// TIA Portal V20 export
Screen "Pop-up_PN_DEV_DIAG_Counter_Popup"  290x322
  ScreenItem "Background" at 0,0 size 290x322  Type=HmiRectangle
  ScreenItem "Text_ReadedDEVNumbers" at 8,163 size 276x25  Type=HmiTextBox
  ScreenItem "Text_Configured" at 10,37 size 130x25  Type=HmiTextBox
  ScreenItem "Counter_Configured" at 145,38 size 44x23  Type=HmiIOField
  ScreenItem "Text_Faulty" at 10,112 size 130x25  Type=HmiTextBox
  ScreenItem "Counter_Faulty" at 145,113 size 44x23  Type=HmiIOField
  ScreenItem "Text_Deaktivated" at 10,87 size 130x25  Type=HmiTextBox
  ScreenItem "Counter_Deaktivated" at 145,88 size 44x23  Type=HmiIOField
  ScreenItem "Text_Present" at 10,62 size 130x25  Type=HmiTextBox
  ScreenItem "Counter_Present" at 145,63 size 44x23  Type=HmiIOField
  ScreenItem "Text_Problem" at 10,137 size 130x25  Type=HmiTextBox
  ScreenItem "Counter_Problem" at 145,138 size 44x23  Type=HmiIOField
  ScreenItem "Text_MaxDevices" at 10,266 size 130x25  Type=HmiTextBox
  ScreenItem "Text_MaxModules" at 10,291 size 130x25  Type=HmiTextBox
  ScreenItem "Counter_MaxDevices" at 145,267 size 44x23  Type=HmiIOField
  ScreenItem "Counter_Max_Modules" at 145,292 size 44x23  Type=HmiIOField
  ScreenItem "Text_PNDEVCounter" at 1,3 size 288x30  Type=HmiTextBox
  ScreenItem "Text_PLCSettings" at 10,241 size 276x25  Type=HmiTextBox
  ScreenItem "Text_Lowest" at 10,185 size 130x25  Type=HmiTextBox
  ScreenItem "Text_Highest" at 10,210 size 130x25  Type=HmiTextBox
  ScreenItem "Counter_LowDevice" at 145,187 size 44x23  Type=HmiIOField
  ScreenItem "Counter_HighDevice" at 145,212 size 44x23  Type=HmiIOField
  ScreenItem "Cancel Mode_1" at 206,278 size 82x42  Type=HmiButton
  ScreenItem "Background_1" at 8,8 size 290x322  Type=HmiRectangle
  ScreenItem "Text_ReadedDEVNumbers_1" at 16,171 size 276x25  Type=HmiTextBox
  ScreenItem "Text_Configured_1" at 18,45 size 130x25  Type=HmiTextBox
  ScreenItem "Counter_Configured_1" at 153,46 size 44x23  Type=HmiIOField
  ScreenItem "Text_Faulty_1" at 18,120 size 130x25  Type=HmiTextBox
  ScreenItem "Counter_Faulty_1" at 153,121 size 44x23  Type=HmiIOField
  ScreenItem "Text_Deaktivated_1" at 18,95 size 130x25  Type=HmiTextBox
  ScreenItem "Counter_Deaktivated_1" at 153,96 size 44x23  Type=HmiIOField
  ScreenItem "Text_Present_1" at 18,70 size 130x25  Type=HmiTextBox
  ScreenItem "Counter_Present_1" at 153,71 size 44x23  Type=HmiIOField
  ScreenItem "Text_Problem_1" at 18,145 size 130x25  Type=HmiTextBox
  ScreenItem "Counter_Problem_1" at 153,146 size 44x23  Type=HmiIOField
  ScreenItem "Text_MaxDevices_1" at 18,274 size 130x25  Type=HmiTextBox
  ScreenItem "Text_MaxModules_1" at 18,299 size 130x25  Type=HmiTextBox
  ScreenItem "Counter_MaxDevices_1" at 153,275 size 44x23  Type=HmiIOField
  ScreenItem "Counter_Max_Modules_1" at 153,300 size 44x23  Type=HmiIOField
  ScreenItem "Text_PNDEVCounter_1" at 9,11 size 288x30  Type=HmiTextBox
  ScreenItem "Text_PLCSettings_1" at 18,249 size 276x25  Type=HmiTextBox
  ScreenItem "Text_Lowest_1" at 18,193 size 130x25  Type=HmiTextBox
  ScreenItem "Text_Highest_1" at 18,218 size 130x25  Type=HmiTextBox
  ScreenItem "Counter_LowDevice_1" at 153,195 size 44x23  Type=HmiIOField
  ScreenItem "Counter_HighDevice_1" at 153,220 size 44x23  Type=HmiIOField
  ScreenItem "Cancel Mode_2" at 214,286 size 82x42  Type=HmiButton
  ScreenItem "Background_2" at 402,11 size 290x322  Type=HmiRectangle
  ScreenItem "Text_ReadedDEVNumbers_2" at 410,174 size 276x25  Type=HmiTextBox
  ScreenItem "Text_Configured_2" at 412,48 size 130x25  Type=HmiTextBox
  ScreenItem "Counter_Configured_2" at 547,49 size 44x23  Type=HmiIOField
  ScreenItem "Text_Faulty_2" at 412,123 size 130x25  Type=HmiTextBox
  ScreenItem "Counter_Faulty_2" at 547,124 size 44x23  Type=HmiIOField
  ScreenItem "Text_Deaktivated_2" at 412,98 size 130x25  Type=HmiTextBox
  ScreenItem "Counter_Deaktivated_2" at 547,99 size 44x23  Type=HmiIOField
  ScreenItem "Text_Present_2" at 412,73 size 130x25  Type=HmiTextBox
  ScreenItem "Counter_Present_2" at 547,74 size 44x23  Type=HmiIOField
  ScreenItem "Text_Problem_2" at 412,148 size 130x25  Type=HmiTextBox
  ScreenItem "Counter_Problem_2" at 547,149 size 44x23  Type=HmiIOField
  ScreenItem "Text_MaxDevices_2" at 412,277 size 130x25  Type=HmiTextBox
  ScreenItem "Text_MaxModules_2" at 412,302 size 130x25  Type=HmiTextBox
  ScreenItem "Counter_MaxDevices_2" at 547,278 size 44x23  Type=HmiIOField
  ScreenItem "Counter_Max_Modules_2" at 547,303 size 44x23  Type=HmiIOField
  ScreenItem "Text_PNDEVCounter_2" at 403,14 size 288x30  Type=HmiTextBox
  ScreenItem "Text_PLCSettings_2" at 412,252 size 276x25  Type=HmiTextBox
  ScreenItem "Text_Lowest_2" at 412,196 size 130x25  Type=HmiTextBox
  ScreenItem "Text_Highest_2" at 412,221 size 130x25  Type=HmiTextBox
  ScreenItem "Counter_LowDevice_2" at 547,198 size 44x23  Type=HmiIOField
  ScreenItem "Counter_HighDevice_2" at 547,223 size 44x23  Type=HmiIOField
  ScreenItem "Cancel Mode_3" at 608,289 size 82x42  Type=HmiButton
